Fanuc KAREL source: kt00903.KL

-- PROVISIONAL review KL for V770-1; original PC SHA256 edab0a9ac97da6e6a2d76b5f9bcf67fa61bba5fbdd4b11347c2b3e42dc1da6c0
-- Incomplete behavior may be omitted. Consult companion uncertainty JSON. Do not deploy.
PROGRAM KT00903
%NOLOCKGROUP
BEGIN
  -- UNRESOLVED_PC offsets 5-28; opcodes 27,22,1C,31,4A
  -- UNRESOLVED_PC offsets 33-37; opcodes 7F
END KT00903
